// TIA Portal V20 export
Screen "PopupAndonLegend"  271x400
  ScreenItem "Text box_30" at 4,20 size 188x24  Type=HmiTextBox
  ScreenItem "Textfeld_Legende" at 13,-1 size 170x25  Type=HmiTextBox
  ScreenItem "Cancel Mode" at 195,3 size 71x42  Type=HmiButton
  ScreenItem "Text box_32" at 4,45 size 188x24  Type=HmiTextBox
  ScreenItem "Text box_33" at 4,70 size 188x24  Type=HmiTextBox
  ScreenItem "Text box_34" at 4,95 size 188x24  Type=HmiTextBox
  ScreenItem "Text box_35" at 4,120 size 188x24  Type=HmiTextBox
  ScreenItem "Text box_36" at 4,145 size 188x24  Type=HmiTextBox
  ScreenItem "Text box_37" at 4,170 size 188x24  Type=HmiTextBox
  ScreenItem "Text box_38" at 4,196 size 188x24  Type=HmiTextBox
  ScreenItem "Text box_39" at 4,221 size 188x24  Type=HmiTextBox
  ScreenItem "Text box_40" at 4,246 size 188x24  Type=HmiTextBox
  ScreenItem "Text box_41" at 4,271 size 188x24  Type=HmiTextBox
  ScreenItem "Text box_42" at 4,296 size 188x24  Type=HmiTextBox
  ScreenItem "Text box_43" at 4,321 size 188x24  Type=HmiTextBox
  ScreenItem "Text box_44" at 4,346 size 188x24  Type=HmiTextBox
  ScreenItem "Text box_45" at 4,372 size 188x24  Type=HmiTextBox
